SUBAPPLICATION GreenWhiteBackground_Abscheider (* Subapplication Type *)
  (* Standard: 61499-2 *)
  (* Version 1.0, 2023-02-06, franz *)
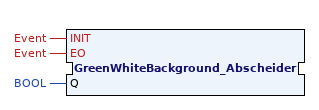
  EVENT_INPUT
    INIT;
    EO;
  END_EVENT
  VAR_INPUT
    Q : BOOL;
  END_VAR
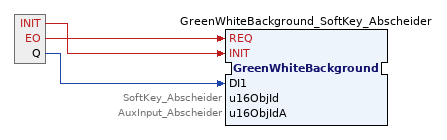
  SUBAPPS
    GreenWhiteBackground_SoftKey_Abscheider : GreenWhiteBackground(u16ObjId := SoftKey_Abscheider, u16ObjIdA := AuxInput_Abscheider);
  END_SUBAPPS
  EVENT_CONNECTIONS
    EO TO GreenWhiteBackground_SoftKey_Abscheider.REQ;
    INIT TO GreenWhiteBackground_SoftKey_Abscheider.INIT;
  END_CONNECTIONS
  DATA_CONNECTIONS
    Q TO GreenWhiteBackground_SoftKey_Abscheider.DI1;
  END_CONNECTIONS
END_SUBAPPLICATION
